(* IEC 61131-3 sources: plc-vscode/tests/st/test-ready/trust-platform/examples/OSCAT/airport_baggage_command_observer/non-oop/src, 3 files *)

(* ---- Main.st ---- *)
FUNCTION_BLOCK ClassicBaggageDiverter
VAR
    LastCommandIdValue : INT;
    EventCountValue : INT;
END_VAR
METHOD PUBLIC ProcessBag : INT
VAR_INPUT
    BagId : INT;
    ScannerResult : INT;
END_VAR
IF ScannerResult = INT#1 THEN
    LastCommandIdValue := INT#1;
ELSIF ScannerResult = INT#2 THEN
    LastCommandIdValue := INT#2;
ELSE
    LastCommandIdValue := INT#3;
END_IF;
EventCountValue := EventCountValue + INT#1;
ProcessBag := LastCommandIdValue;
END_METHOD
PUBLIC PROPERTY EventCount : INT
GET
    EventCount := EventCountValue;
END_GET
END_PROPERTY
END_FUNCTION_BLOCK
PROGRAM Main
VAR
    Diverter : ClassicBaggageDiverter;
    Command : INT;
END_VAR
Command := Diverter.ProcessBag(BagId := INT#42, ScannerResult := INT#2);
END_PROGRAM

(* ---- Configuration.st ---- *)
CONFIGURATION AirportBaggageCommandObserverClassicConfiguration
RESOURCE Cpu0 ON PLC
    TASK MainTask (INTERVAL := T#50ms, PRIORITY := 1);
    PROGRAM Diverter WITH MainTask : Main;
END_RESOURCE
END_CONFIGURATION

(* ---- Tests.st ---- *)
TEST_PROGRAM ClassicBaggageBranchesOnScannerResult
VAR
    Diverter : ClassicBaggageDiverter;
END_VAR
ASSERT_EQUAL(EXPECTED := INT#2, ACTUAL := Diverter.ProcessBag(BagId := INT#42, ScannerResult := INT#2));
ASSERT_EQUAL(EXPECTED := INT#1, ACTUAL := Diverter.EventCount);
END_TEST_PROGRAM
